(* IEC 61131-3 sources: plc-iiot-stack/src/POUs/Iiot/F_IiotCmdFromString, 2 files *)

(* ---- F_IiotCmdFromString.decl.st ---- *)
// Назначение: команда по имени поля command (с учётом регистра, enum command.schema.json);
//             неизвестное имя — None.
// Автор:      kr0nsch
// Версия:     0.1.0
// Документ:   docs/plc_mqtt.md, раздел «Команды»
FUNCTION F_IiotCmdFromString : E_IiotCommand
VAR_INPUT
    sCommand : STRING(GVL_Const.JSON_STR_LEN);
END_VAR

(* ---- F_IiotCmdFromString.impl.st ---- *)
IF sCommand = 'SetAuto' THEN
    F_IiotCmdFromString := E_IiotCommand.SetAuto;
ELSIF sCommand = 'SetManual' THEN
    F_IiotCmdFromString := E_IiotCommand.SetManual;
ELSIF sCommand = 'SetOos' THEN
    F_IiotCmdFromString := E_IiotCommand.SetOos;
ELSIF sCommand = 'Start' THEN
    F_IiotCmdFromString := E_IiotCommand.Start;
ELSIF sCommand = 'Stop' THEN
    F_IiotCmdFromString := E_IiotCommand.Stop;
ELSIF sCommand = 'SpeedSp' THEN
    F_IiotCmdFromString := E_IiotCommand.SpeedSp;
ELSIF sCommand = 'ResetMaint' THEN
    F_IiotCmdFromString := E_IiotCommand.ResetMaint;
ELSIF sCommand = 'SubstValue' THEN
    F_IiotCmdFromString := E_IiotCommand.SubstValue;
ELSIF sCommand = 'Ack' THEN
    F_IiotCmdFromString := E_IiotCommand.Ack;
ELSIF sCommand = 'Reset' THEN
    F_IiotCmdFromString := E_IiotCommand.Reset;
ELSIF sCommand = 'AckReq' THEN
    F_IiotCmdFromString := E_IiotCommand.AckReq;
ELSIF sCommand = 'ShelveReq' THEN
    F_IiotCmdFromString := E_IiotCommand.ShelveReq;
ELSIF sCommand = 'UnshelveReq' THEN
    F_IiotCmdFromString := E_IiotCommand.UnshelveReq;
ELSIF sCommand = 'SetStepped' THEN
    F_IiotCmdFromString := E_IiotCommand.SetStepped;
ELSIF sCommand = 'SetLevelPid' THEN
    F_IiotCmdFromString := E_IiotCommand.SetLevelPid;
ELSIF sCommand = 'AckAll' THEN
    F_IiotCmdFromString := E_IiotCommand.AckAll;
ELSIF sCommand = 'ResetAll' THEN
    F_IiotCmdFromString := E_IiotCommand.ResetAll;
ELSIF sCommand = 'Silence' THEN
    F_IiotCmdFromString := E_IiotCommand.Silence;
ELSE
    F_IiotCmdFromString := E_IiotCommand.None;
END_IF
